Fanuc KAREL source: kb00079.KL

PROGRAM KB00079
%STACKSIZE=65535
%PRIORITY=65535
%NOLOCKGROUP
VAR
P1 : INTEGER
P2 : INTEGER
P3 : INTEGER
RESULT : JOINTPOS9
BEGIN
P1=1
P2=1
P3=1
-- UNSAFE_SOURCE_IR line 12: CALL_RESULT GET_JPOS_TPE(P1, P2, P3, 1)
END KB00079
